Fanuc KAREL source: KB00194.KL

PROGRAM KB00194
%NOLOCKGROUP
VAR
  P1: STRING[80]
  P2: INTEGER
  P3: INTEGER
BEGIN
  P1 = 'A'
  P2 = 1
  P3 = 1
  V_GET_OFFSET(P1, P2, P3)
END KB00194
